// TIA Portal V21 export
// export: Created 2026-11-08T21:17:25.6740455Z, ExportSetting WithDefaults, DisplayName Totally Integrated Automation Portal, DisplayVersion V21 Update 3, DisplayName STEP 7 Professional, DisplayVersion V21 Update 3, DisplayName STEP 7 Safety, DisplayVersion V21, DisplayName Tech WebApplication, DisplayVersion V21, DisplayName WinCC Basic/Comfort/Advanced, DisplayVersion V21 Update 3, DisplayName WinCC Unified, DisplayVersion V21 Update 3
DATA_BLOCK "FB_Iface_DB"   // DB5
VERSION : 0.1
// stored: AutoNumber true, DBAccessibleFromOPCUA true, DBAccessibleFromWebserver true, InstanceOfName FB_Iface, InstanceOfType FB
"FB_Iface"
   // VAR_INPUT
   //    iBool : Bool;
   //    iInt : Int;
   //    iReal : Real;
   //    iArr : Array[0..3] of Int;
   //    iMotor : "UDT_Motor";
   // END_VAR
   // VAR_OUTPUT
   //    oBool : Bool;
   //    oInt : Int;
   // END_VAR
   // VAR_IN_OUT
   //    ioReal : Real;
   // END_VAR
   // VAR
   //    stInt : Int := 99;
   //    stBool : Bool := TRUE;
   // END_VAR
BEGIN
END_DATA_BLOCK
